DATA_BLOCK "FRK_Views"
{ S7_Optimized_Access := 'TRUE' }
VERSION : 0.1
NON_RETAIN
VAR
    V001 {ExternalAccessible := 'False'; ExternalVisible := 'False'; ExternalWritable := 'False'} : "FRK_ViewOwned_DeclarationUnit";
    V013 {ExternalAccessible := 'False'; ExternalVisible := 'False'; ExternalWritable := 'False'} : "FRK_ViewOwned_DeclarationUnit";
END_VAR
BEGIN
END_DATA_BLOCK
